(*
SPDX-FileCopyrightText: © 2026 Oleksandr Tiutyk <trofimich@gmail.com>
SPDX-License-Identifier: MIT
License: https://opensource.org/license/mit
*)

(*!
<summary>Waits until a configured workflow condition evaluates to TRUE.</summary>
<description>
Evaluates the attached condition cyclically in ACTIVE_RUNNING. Transitions to PASSIVE_COMPLETED when the
condition returns TRUE. Cancelling or suspending stops waiting immediately.
</description>
*)

{attribute 'no_explicit_call' := 'do not call this function block directly'}
{attribute 'enable_dynamic_creation'}
FUNCTION_BLOCK WaitConditionActivity EXTENDS Activity
	IMPLEMENTS IWaitConditionActivity, TOF_Core.IConfigurationSerializable
VAR_STAT
	{attribute 'hide'}
	_ClassName : STRING := __POUNAME();
END_VAR
VAR
	{attribute 'OPC.UA.DA' := '0'}
	_Condition : ICondition;

	{attribute 'OPC.UA.DA' := '0'}
	_Configured : BOOL;
END_VAR

(*!
<summary>Borrows the initialized class name used in diagnostics.</summary>
<description>
Returns initialized metadata storage without allocation. Callers must not modify the returned string.
Derived function blocks must use distinct initialized static storage when overriding this metadata.
</description>
*)
{attribute 'monitoring' := 'call'}
PROPERTY ClassName : REFERENCE TO STRING
GET
ClassName REF= _ClassName;
END_GET
END_PROPERTY

(*!
<summary>Returns the condition being evaluated, or 0 before configuration.</summary>
*)
{attribute 'monitoring' := 'call'}
PROPERTY Condition : ICondition
GET
Condition := _Condition;
END_GET
END_PROPERTY

(*!
<summary>Configures the condition to wait for.</summary>
<description>
Validates that the condition is live, unattached to another parent, and establishes the parent link.
The parent chain and owning workflow must be PASSIVE_READY; fixed workflow association is checked before
mutation. Reusing the same dependency is permitted. Replaced dependencies retain their existing parent links
and must not be attached elsewhere. Parent callbacks are not transactional. Dependencies remain borrowed.
</description>
<param name="condition">Condition to evaluate during execution.</param>
*)
METHOD Configure
VAR_INPUT
	condition : ICondition;
END_VAR
IF condition = 0 THEN
	TOF_Core.Exceptions.ThrowArgumentNotSpecified(
		sourceNamespaceName := NamespaceName,
		sourceClassName := ClassName,
		sourcePOUName := __POUNAME(),
		sourcePosition := __POSITION(),
		argumentName := 'condition'
	);
END_IF

Workflows.ValidateElementAttachment(parent := THIS^, child := condition);

_Configured := FALSE;

_Condition := condition;
_Condition.ParentActivity := THIS^;

_Configured := TRUE;
END_METHOD

(*!
<summary>Reports whether the condition has been configured.</summary>
*)
{attribute 'monitoring' := 'call'}
PROPERTY Configured : BOOL
GET
Configured := _Configured;
END_GET
END_PROPERTY

(*!
<summary>Borrows the compiler-initialized library namespace.</summary>
<description>
Borrows storage from the live internal namespace provider. Reacquire references after application
reinitialization or relocation. Treat the reference as read-only; no ownership or synchronization is provided.
</description>
*)
{attribute 'monitoring' := 'call'}
PROPERTY NamespaceName : REFERENCE TO STRING
GET
NamespaceName REF= CurrentNamespace.Name;
END_GET
END_PROPERTY

(*!
<summary>Completes resetting in a single step.</summary>
<param name="startResetting">TRUE on the initial call from RequestReset.</param>
*)
METHOD PROTECTED OnResetting : ACTIVITY_RESETTING_STATE
VAR_INPUT
	startResetting : BOOL;
END_VAR
OnResetting := ACTIVITY_RESETTING_STATE.WORK_RESET;
END_METHOD

(*!
<summary>Evaluates the configured condition and completes when it returns TRUE.</summary>
<param name="startRunning">TRUE on the initial call of a fresh start.</param>
<param name="startResuming">TRUE when resuming execution after suspension.</param>
<param name="haltReason">Unused halt reason output.</param>
*)
METHOD PROTECTED OnRunning : ACTIVITY_RUNNING_STATE
VAR_INPUT
	startRunning : BOOL;
	startResuming : BOOL;
END_VAR
VAR_OUTPUT
	haltReason : WSTRING(255);
END_VAR
IF NOT _Configured THEN
	WorkflowExceptions.ThrowWorkflowConfiguration(
		sourceNamespaceName := NamespaceName,
		sourceClassName := ClassName,
		sourcePOUName := __POUNAME(),
		sourcePosition := __POSITION(),
		message := "Activity is not configured"
	);
END_IF

IF _Condition.Evaluate(activity := THIS^) THEN
	OnRunning := ACTIVITY_RUNNING_STATE.WORK_COMPLETED;
END_IF
END_METHOD

(*!
<summary>Stops waiting immediately on cancel or suspend.</summary>
<param name="startCancelling">TRUE when stopping due to cancellation.</param>
<param name="startSuspending">TRUE when stopping due to suspension.</param>
<param name="haltReason">Unused halt reason output.</param>
*)
METHOD PROTECTED OnStopping : ACTIVITY_STOPPING_STATE
VAR_INPUT
	startCancelling : BOOL;
	startSuspending : BOOL;
END_VAR
VAR_OUTPUT
	haltReason : WSTRING(255);
END_VAR
OnStopping := ACTIVITY_STOPPING_STATE.WORK_STOPPED;
END_METHOD

(*!
<summary>Reports the size of this concrete function block instance in bytes.</summary>
<description>
Reports the instance layout rather than dynamic allocations owned by its fields. A derived function block
with a different layout must override this property; the value does not grant disposal rights.
</description>
*)
{attribute 'monitoring' := 'call'}
PROPERTY SelfSize : ULINT
GET
SelfSize := XSIZEOF(THIS^);
END_GET
END_PROPERTY

(*!
<summary>Writes the configuration fields for this object.</summary>
<description>Borrows the writer for this call. A failure invalidates the current output document.</description>
*)
METHOD Serialize
VAR_INPUT
	writer : TOF_Core.IConfigurationWriter;
END_VAR
Workflows.WriteConfigurationHeader(writer := writer, source := THIS^, displayName := Name, scope := THIS^);
Workflows.WriteConfigurationObject(writer := writer, name := 'condition', source := _Condition);
END_METHOD

(*!
<summary>Restores this fresh instance from its configuration object.</summary>
<description>
The reader, document node and deserialization context are borrowed for this call.
On failure discard the partial instance.
</description>
<param name="reader">Active configuration reader.</param>
<param name="node">Object node to read fields from.</param>
<param name="context">Active configuration deserialization context providing workflow reconstruction services.</param>
*)
METHOD Deserialize
VAR_INPUT
	reader : TOF_Core.IConfigurationReader;
	node : TOF_Core.CONFIGURATION_NODE;
	context : TOF_Core.IConfigurationDeserializationContext;
END_VAR
VAR
	loader : IWorkflowLoader;
END_VAR
loader := WorkflowConfigurationSerializer.ResolveWorkflowLoader(context := context);
Workflows.ReadConfigurationHeader(reader := reader, node := node, target := THIS^, scope := THIS^);

Configure(
	condition := Workflows.ReadCondition(
		loader := loader,
		node := reader.GetField(node := node, name := 'condition')
	)
);
END_METHOD

END_FUNCTION_BLOCK

(* stored: Version 1.1.0.1
   POU WaitConditionActivity: Id {0916704d-d918-47c7-8c0e-c8da18f42f13}, SpecialFunc None
   Folder Overriden methods: Id {88b71d49-47c0-482a-a9e1-253198de7401}
   Property ClassName: Id {d1752f9e-57cf-4764-a0c1-9ed82f64081e}
   Get Get: Id {0142adec-9a1f-40ba-9edf-55dab0af9cb3}
   Property Condition: Id {09cb088a-beaf-41db-a5bb-81751b0a87ab}
   Get Get: Id {ebfbe611-3ed2-4287-9d89-a3a34c1b445d}
   Method Configure: Id {52e11014-c0d9-473e-a276-5438377e75e8}
   Property Configured: Id {c0b002fa-3d61-4b93-ac3e-bed6aec10d4a}
   Get Get: Id {8764b566-fd9f-4d8f-b740-bcb39bd3ca7a}
   Property NamespaceName: Id {d2aa2dd8-7c8d-4c49-a66c-eb757eb24965}
   Get Get: Id {42870797-7f65-46e6-84e4-80b3ea493422}
   Method OnResetting: Id {4e25309c-9bda-4398-8979-3f8c64d201d2}
   Method OnRunning: Id {f56a370a-0201-439d-b79b-b4a23784d2df}
   Method OnStopping: Id {7d8c16f6-b73b-4b3e-b96f-ccd88ad1a7d4}
   Property SelfSize: Id {17ad9913-b398-4404-a687-463af48f4ef4}
   Get Get: Id {9029c1e2-7d7d-492d-b7b0-360bebbc6748}
   Method Serialize: Id {0b07211a-d2a8-4cce-8346-290d53ff080e}
   Method Deserialize: Id {bbc96361-3dd1-48ff-b9fb-542bb0f542d2} *)
